// Mitsubishi GX Works2 project: 타이머+모터   PLC: Q02/Q02H

PROGRAM MAIN
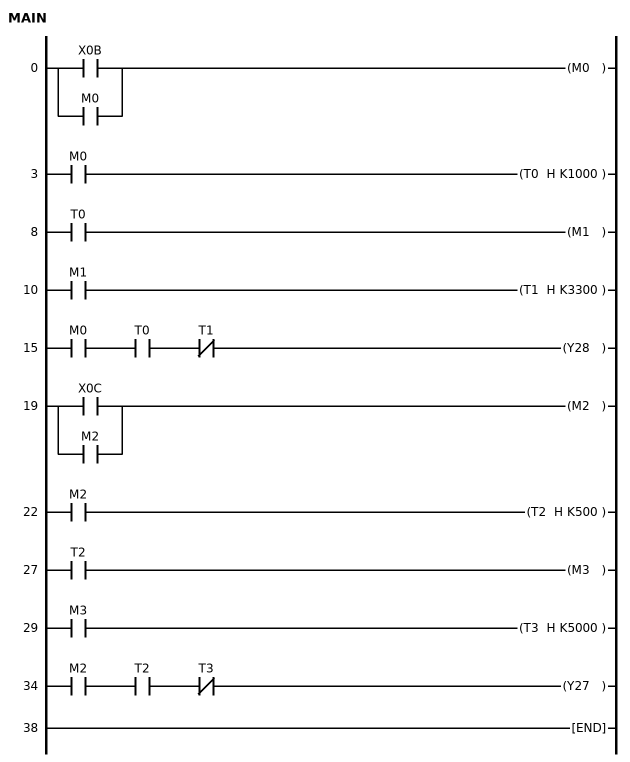
0     LD      X0B
      OR      M0
      OUT     M0
3     LD      M0
      OUTH    T0 K1000
8     LD      T0
      OUT     M1
10    LD      M1
      OUTH    T1 K3300
15    LD      M0
      AND     T0
      ANI     T1
      OUT     Y28
19    LD      X0C
      OR      M2
      OUT     M2
22    LD      M2
      OUTH    T2 K500
27    LD      T2
      OUT     M3
29    LD      M3
      OUTH    T3 K5000
34    LD      M2
      AND     T2
      ANI     T3
      OUT     Y27
38    END
END_PROGRAM
